(* IEC 61131-3 sources: s22-soft-shell/st_interpret/tests/test_inputs/st_stretch, 1 file *)

(* ---- stretch_pow.st ---- *)
PROGRAM stretch_pow
VAR
    a: int;
END_VAR
    a := 3 ** 3;
END_PROGRAM
